Fanuc KAREL source: kt00483.KL

-- PROVISIONAL review KL for V1013-1; original PC SHA256 c2f05d5c4007e0ed382c99dfa8f565c46ac3e1f8e22d739b457d5d161c59ad54
-- Incomplete behavior may be omitted. Consult companion uncertainty JSON. Do not deploy.
PROGRAM KT00483
%NOLOCKGROUP
VAR
  OUT : BOOLEAN
-- UNRESOLVED_DECL P1 type=000101
-- UNRESOLVED_DECL P2 type=000106
BEGIN
  -- UNRESOLVED_PC offsets 5-20; opcodes 2E,22,32,35
  -- UNRESOLVED_PC offsets 25-53; opcodes 49,49,7E,AC,23
  -- UNRESOLVED_PC offsets 58-62; opcodes 7F
END KT00483
